Fanuc KAREL source: kc00003.KL

-- PROVISIONAL review KL for V940-1; original PC SHA256 93859522449f1cf32e990df60fbe35a94d3567e342ade452aa06f262bcb964e8
-- Incomplete behavior may be omitted. Consult companion uncertainty JSON. Do not deploy.
PROGRAM KC00003
%NOLOCKGROUP
BEGIN
  -- V9_ZERO_TABLE_METADATA_HINT layout=0002_ascii; no indexed target words; source/name/runtime held
  -- UNRESOLVED_PC offsets 5-33; opcodes 27,22,22,22,22,31
  -- UNRESOLVED_PC offsets 38-42; opcodes 7F
END KC00003
